Fanuc KAREL source: KO00063.KL

PROGRAM KO00063
%NOLOCKGROUP
%ENVIRONMENT MIR
VAR
  P1: XYZWPR
  P2: JOINTPOS
  F: BOOLEAN
  OUT: XYZWPREXT
BEGIN
  F = TRUE
  OUT = MIRROR(P1, P2, F)
END KO00063
